(* IEC 61131-3 sources: llm-plc-st-eval/codesys (part 2) *)

(* ---- PRG_Test_I2.st ---- *)
(*
    BANCO DE PRUEBA AUTOVERIFICABLE — Tarea I2 (FSM de llenado multietapa)
    ---------------------------------------------------------------------------
    Reposo -> llenado -> mezcla 60 s -> descarga -> reposo. El paro debe llevar
    a estado seguro (todas las salidas desactivadas) desde CUALQUIER etapa y
    devolver el proceso a reposo.

    USO: crear este PROGRAM junto al FUNCTION_BLOCK de la respuesta a evaluar y
    ejecutar en modo Simulacion. Al terminar, leer 'veredicto': 1 = supera,
    2 = falla.

    ---------------------------------------------------------------------------
    CORRECCION DEL 2026-09-09 (enmienda 10). Validado con validar_harness_I2.py.
    La version anterior tenia dos fallos:

    FALLO 1 — el paso de "antes de los 60 s" REPROBABA a la implementacion
    correcta en los tres ciclos de tarea. Esperaba 59 800 ms contando desde el
    inicio de ese paso, pero la mezcla no arranca ahi: arranca ~200 ms antes,
    en el paso anterior, en cuanto el bloque ve nivelAlto. El margen resultante
    era nulo y la evaluacion caia justo en el instante en que la mezcla
    termina, de modo que se observaba ya la descarga. Es el mismo error que la
    enmienda 5 corrigio en I4: una ventana calculada como si la fase empezara
    en el limite del paso, cuando empieza antes.

    FALLO 2 — el ultimo paso, etiquetado "paro en mezcla", NUNCA llegaba a la
    mezcla. Aplicaba nivelAlto y btnParo en el MISMO paso, asi que el paro
    alcanzaba al bloque todavia en llenado: era un duplicado del paso anterior.
    Verificado: una implementacion cuyo paro funciona en llenado pero no
    durante la mezcla obtenia el mismo resultado que la correcta. El paro en
    dos fases que este banco dice comprobar solo se comprobaba en una.

    La correccion de tiempos de este documento ya lo insinuaba al estimar I2 en
    ~90 s "porque el paro se prueba en dos fases distintas, cada una exige
    volver a entrar en la fase": la secuencia real duraba 61,9 s porque esa
    segunda entrada nunca se hacia.

    Correcciones: la ventana de la mezcla pasa a tener margen explicito y
    simetrico de 0,5 s a cada lado de los 60 s; y entrar en la mezcla y aplicar
    el paro pasan a ser dos pasos separados, de modo que el paro alcance al
    bloque realmente mezclando. Se anade ademas un paso final que comprueba que
    tras el paro el proceso permanece en reposo y no rearranca solo.
*)

PROGRAM PRG_Test_I2
VAR CONSTANT
    ULTIMO_PASO : INT := 11;          (* 12 pasos: indices 0..11 *)
END_VAR
VAR
    (* --- Bloque bajo prueba: sustituir por la respuesta a evaluar --- *)
    fb : FB_Llenado;

    (* --- Entradas manipuladas por el banco --- *)
    nivelAlto : BOOL;
    nivelBajo : BOOL;
    btnInicio : BOOL;
    btnParo   : BOOL;

    (* --- Control de la secuencia --- *)
    evL, evM, evD : BOOL;
    paso       : INT := 0;
    tEspera    : TIME;
    tPaso      : TON;
    pulsoReset : BOOL;
    finalizado : BOOL;

    (* --- Resultados: 0 = pendiente, 1 = pasa, 2 = falla --- *)
    resultado : ARRAY[0..11] OF INT;
    nPasan    : INT;
    veredicto : INT := 0;
    i         : INT;
END_VAR

(* 1. Definicion del paso en curso *)
IF NOT finalizado THEN
    CASE paso OF
        0:  (* Reposo *)
            nivelAlto := FALSE; nivelBajo := FALSE;
            btnInicio := FALSE; btnParo := FALSE;
            tEspera := T#200MS; evL := FALSE; evM := FALSE; evD := FALSE;
        1:  (* Arranque: abre la valvula de llenado *)
            btnInicio := TRUE;
            tEspera := T#200MS; evL := TRUE;  evM := FALSE; evD := FALSE;
        2:  (* Nivel alto: entra en mezcla. La mezcla arranca AQUI, no en el
               paso siguiente; de ahi el margen explicito del paso 3. *)
            btnInicio := FALSE; nivelAlto := TRUE;
            tEspera := T#1S;    evL := FALSE; evM := TRUE;  evD := FALSE;
        3:  (* ~59,5 s de mezcla acumulados: aun NO debe haber terminado *)
            tEspera := T#58500MS; evM := TRUE;
        4:  (* ~60,5 s acumulados: ya debe estar descargando *)
            tEspera := T#1S;    evL := FALSE; evM := FALSE; evD := TRUE;
        5:  (* Nivel bajo: vuelve a reposo *)
            nivelBajo := TRUE;
            tEspera := T#200MS; evL := FALSE; evM := FALSE; evD := FALSE;

        (* --- Paro en la fase de LLENADO --- *)
        6:  (* Nuevo ciclo *)
            nivelAlto := FALSE; nivelBajo := FALSE; btnInicio := TRUE;
            tEspera := T#200MS; evL := TRUE;  evM := FALSE; evD := FALSE;
        7:  (* Paro estando en llenado: estado seguro *)
            btnInicio := FALSE; btnParo := TRUE;
            tEspera := T#200MS; evL := FALSE; evM := FALSE; evD := FALSE;

        (* --- Paro en la fase de MEZCLA (enmienda 10): entrar en la mezcla y
               aplicar el paro son DOS pasos distintos, para que el paro
               alcance al bloque realmente mezclando --- *)
        8:  (* Rearranca tras el paro *)
            btnParo := FALSE; btnInicio := TRUE;
            tEspera := T#200MS; evL := TRUE;  evM := FALSE; evD := FALSE;
        9:  (* Entra en mezcla y se deja mezclando *)
            btnInicio := FALSE; nivelAlto := TRUE;
            tEspera := T#500MS; evL := FALSE; evM := TRUE;  evD := FALSE;
        10: (* Paro ESTANDO EN MEZCLA: estado seguro *)
            btnParo := TRUE;
            tEspera := T#200MS; evL := FALSE; evM := FALSE; evD := FALSE;
        11: (* Tras el paro debe permanecer en reposo, sin rearrancar solo *)
            btnParo := FALSE; nivelAlto := FALSE;
            tEspera := T#200MS; evL := FALSE; evM := FALSE; evD := FALSE;
    END_CASE
END_IF

(* 2. Temporizador de asentamiento del paso *)
tPaso(IN := NOT pulsoReset, PT := tEspera);
pulsoReset := FALSE;

(* 3. Llamada al bloque bajo prueba *)
fb(nivelAlto := nivelAlto, nivelBajo := nivelBajo,
   btnInicio := btnInicio, btnParo := btnParo);

(* 4. Evaluacion al vencer el asentamiento *)
IF tPaso.Q AND NOT finalizado THEN
    IF fb.vLlenado = evL AND fb.motorMezcla = evM AND fb.vDescarga = evD THEN
        resultado[paso] := 1;
    ELSE
        resultado[paso] := 2;
    END_IF

    pulsoReset := TRUE;

    IF paso < ULTIMO_PASO THEN
        paso := paso + 1;
    ELSE
        finalizado := TRUE;
    END_IF
END_IF

(* 5. Veredicto global *)
IF finalizado AND veredicto = 0 THEN
    nPasan := 0;
    FOR i := 0 TO ULTIMO_PASO DO
        IF resultado[i] = 1 THEN
            nPasan := nPasan + 1;
        END_IF
    END_FOR

    IF nPasan = (ULTIMO_PASO + 1) THEN
        veredicto := 1;
    ELSE
        veredicto := 2;
    END_IF
END_IF

(* ---- PRG_Test_I3.st ---- *)
(*
    BANCO DE PRUEBA AUTOVERIFICABLE — Tarea I3 (gestion de alarmas con prioridad)
    ---------------------------------------------------------------------------
    Tres alarmas con prioridad (alm1 alta, alm2 media, alm3 baja). Cualquiera
    activa enciende la sirena. codigoAlm reporta la de mayor prioridad presente
    (0 si no hay). Cada alarma queda RETENIDA aunque su causa desaparezca hasta
    que se reconozca individualmente, y el reconocimiento SOLO tiene efecto si
    la causa ya desaparecio.

    USO: crear este PROGRAM junto al FUNCTION_BLOCK de la respuesta a evaluar y
    ejecutar en modo Simulacion. Al terminar, leer 'veredicto': 1 = supera,
    2 = falla.

    ---------------------------------------------------------------------------
    CORRECCION DEL 2026-09-09 (enmienda 12). Validado con validar_harness_I3.py.
    La version anterior daba veredicto 1 a una implementacion cuyo ACK borraba
    la alarma AUNQUE la causa siguiera presente, que es la violacion directa de
    la regla central del enunciado. Los nueve pasos daban exactamente el mismo
    resultado que con la implementacion correcta.

    Causa: en toda la secuencia no habia un solo instante en que una entrada
    ackN estuviera activa a la vez que su almN. Los reconocimientos se
    aplicaban siempre con la causa ya retirada, de modo que la mitad de la
    regla ("no debe borrar con la causa presente") no se ejercitaba nunca.

    Es notable porque ENMIENDAS_HARNESSES.md ya aprobaba explicitamente ese
    paso en su lista: "I3: ACK con la causa todavia presente (no debe borrar) y
    ACK tras retirarla (si debe)". El paso estaba aprobado en el documento pero
    no implementado en el banco.

    Correccion: se anade el paso 2, que aplica ack3 con alm3 todavia activa y
    exige que la alarma NO se borre. La secuencia pasa de 9 a 10 pasos.
*)

PROGRAM PRG_Test_I3
VAR CONSTANT
    ULTIMO_PASO    : INT  := 9;       (* 10 pasos: indices 0..9 *)
    T_ASENTAMIENTO : TIME := T#150MS;
END_VAR
VAR
    (* --- Bloque bajo prueba: sustituir por la respuesta a evaluar --- *)
    fb : FB_Alarmas;

    (* --- Entradas manipuladas por el banco --- *)
    alm1, alm2, alm3 : BOOL;
    ack1, ack2, ack3 : BOOL;

    (* --- Control de la secuencia --- *)
    espSirena  : BOOL;
    espCodigo  : INT;
    paso       : INT := 0;
    tPaso      : TON;
    pulsoReset : BOOL;
    finalizado : BOOL;

    (* --- Resultados: 0 = pendiente, 1 = pasa, 2 = falla --- *)
    resultado : ARRAY[0..9] OF INT;
    nPasan    : INT;
    veredicto : INT := 0;
    i         : INT;
END_VAR

(* 1. Temporizador de asentamiento entre pasos *)
tPaso(IN := NOT pulsoReset, PT := T_ASENTAMIENTO);
pulsoReset := FALSE;

(* 2. Aplicacion de entradas y valores esperados. Solo se asigna lo que cada
      paso cambia: las demas entradas conservan su valor. *)
IF NOT finalizado THEN
    CASE paso OF
        0:  (* Reposo: sin alarmas, con los ACK activos (no deben hacer nada) *)
            alm1 := FALSE; alm2 := FALSE; alm3 := FALSE;
            ack1 := TRUE;  ack2 := TRUE;  ack3 := TRUE;
            espSirena := FALSE; espCodigo := 0;
        1:  (* Alarma baja activa *)
            ack1 := FALSE; ack2 := FALSE; ack3 := FALSE;
            alm3 := TRUE;
            espSirena := TRUE;  espCodigo := 3;
        2:  (* ACK CON LA CAUSA TODAVIA PRESENTE: no debe borrar (enmienda 12) *)
            ack3 := TRUE;
            espSirena := TRUE;  espCodigo := 3;
        3:  (* Se retira la causa y se suelta el ACK: sigue retenida *)
            alm3 := FALSE; ack3 := FALSE;
            espSirena := TRUE;  espCodigo := 3;
        4:  (* ACK con la causa ya retirada: ahora si debe borrar *)
            ack3 := TRUE;
            espSirena := FALSE; espCodigo := 0;
        5:  (* Dos alarmas: domina la de mayor prioridad de las presentes *)
            ack3 := FALSE; alm2 := TRUE; alm3 := TRUE;
            espSirena := TRUE;  espCodigo := 2;
        6:  (* Entra la de prioridad alta *)
            alm1 := TRUE;
            espSirena := TRUE;  espCodigo := 1;
        7:  (* Se retira y reconoce la alta: queda la media *)
            alm1 := FALSE; ack1 := TRUE;
            espSirena := TRUE;  espCodigo := 2;
        8:  (* Se retira y reconoce la media: queda la baja *)
            alm2 := FALSE; ack2 := TRUE;
            espSirena := TRUE;  espCodigo := 3;
        9:  (* Se retira y reconoce la baja: todo en reposo *)
            alm3 := FALSE; ack3 := TRUE;
            espSirena := FALSE; espCodigo := 0;
    END_CASE
END_IF

(* 3. Llamada al bloque bajo prueba *)
fb(alm1 := alm1, alm2 := alm2, alm3 := alm3,
   ack1 := ack1, ack2 := ack2, ack3 := ack3);

(* 4. Evaluacion al vencer el asentamiento *)
IF tPaso.Q AND NOT finalizado THEN
    IF fb.sirena = espSirena AND fb.codigoAlm = espCodigo THEN
        resultado[paso] := 1;
    ELSE
        resultado[paso] := 2;
    END_IF

    pulsoReset := TRUE;

    IF paso < ULTIMO_PASO THEN
        paso := paso + 1;
    ELSE
        finalizado := TRUE;
    END_IF
END_IF

(* 5. Veredicto global *)
IF finalizado AND veredicto = 0 THEN
    nPasan := 0;
    FOR i := 0 TO ULTIMO_PASO DO
        IF resultado[i] = 1 THEN
            nPasan := nPasan + 1;
        END_IF
    END_FOR

    IF nPasan = (ULTIMO_PASO + 1) THEN
        veredicto := 1;
    ELSE
        veredicto := 2;
    END_IF
END_IF

(* ---- PRG_Test_I4.st ---- *)
(*
    BANCO DE PRUEBA AUTOVERIFICABLE — Tarea I4 (arranque estrella-triangulo)
    ---------------------------------------------------------------------------
    Aplica la enmienda 2 de ENMIENDAS_HARNESSES.md: DOS verificaciones
    independientes, porque una transicion con 0 ms de tiempo muerto no produce
    ningun scan con kY AND kD y por tanto la bandera de interlock por si sola
    no la detecta.
      1. Seguridad (continua y enclavada): si en cualquier scan kY AND kD, la
         bandera 'interlock' queda en TRUE hasta el final del banco.
      2. Tiempo muerto (medido): se cronometra el intervalo entre la caida de
         kY y la subida de kD y se exige que alcance el minimo.

    Ciclo de MainTask: 4 a 10 ms (enmienda 3). El umbral del tiempo muerto
    absorbe un ciclo de cuantizacion del scan.

    USO: crear este PROGRAM junto al FUNCTION_BLOCK de la respuesta a evaluar y
    ejecutar en modo Simulacion. Al terminar, leer 'veredicto': 1 = supera,
    2 = falla. 'resultado' indica el paso; 'interlock' y 'duracionMuerto' se
    registran aparte porque una violacion de seguridad es cualitativamente
    distinta de un fallo funcional (enmienda 4).

    ---------------------------------------------------------------------------
    CORRECCION DEL 2026-09-09 (enmienda 5). La version anterior tenia tres
    fallos, verificados por simulacion con validar_harness_I4.py:

      1. El paso 2 exigia NOT kD a los 8,3 s, cuando una implementacion
         correcta ya tiene el triangulo dentro desde los 8,1 s. Reprobaba al
         100 % de las implementaciones validas. Era un residuo del enfoque de
         muestreo que la enmienda 2 habia descartado.
      2. La medida reiniciaba su temporizador con un ciclo de retraso, de modo
         que contaba de menos alrededor de un scan: un tiempo muerto correcto
         de 100 ms se media como 96 ms con ciclo de 4 ms y 80 ms con 20 ms, y
         se comparaba contra un umbral estricto de 100 ms.
      3. Si kY caia y kD subia en el MISMO scan, ambas condiciones se cumplian
         en el mismo ciclo, la medida leia un valor viejo del cronometro y
         registraba 8 208 ms: daba por bueno el defecto de 0 ms de tiempo
         muerto, que es exactamente el que la enmienda 2 persigue.

    La medida pasa a hacerse por DIFERENCIA de dos lecturas de un cronometro
    libre que nunca se reinicia. Eso elimina el retraso de un ciclo y hace que
    el caso simultaneo mida 0 ms por construccion, sin necesidad de un caso
    especial. El paso 2 pasa a comprobar que la transicion se completo, y el
    instante exacto queda a cargo de la medida en el paso 3.
*)

PROGRAM PRG_Test_I4
VAR CONSTANT
    ULTIMO_PASO   : INT  := 5;
    T_MUERTO_MIN  : TIME := T#90MS;   (* 100 ms del enunciado menos un ciclo de
                                         MainTask: la cuantizacion del scan es
                                         inevitable y se declara en la metodologia *)
    T_CRONO       : TIME := T#100S;   (* cronometro libre: nunca se reinicia *)
END_VAR
VAR
    (* --- Bloque bajo prueba: sustituir por la respuesta a evaluar --- *)
    fb : FB_EstrellaTriangulo;

    (* --- Entradas manipuladas por el banco --- *)
    btnMarcha : BOOL;
    btnParo   : BOOL;

    (* --- Control de la secuencia --- *)
    paso       : INT := 0;
    tEspera    : TIME;
    tPaso      : TON;
    pulsoReset : BOOL;
    finalizado : BOOL;

    (* --- Verificacion 1: seguridad continua y enclavada (enmiendas 2 y 4) --- *)
    interlock : BOOL;

    (* --- Verificacion 2: medida del tiempo muerto (enmienda 2) --- *)
    tCrono         : TON;
    prevY, prevD   : BOOL;
    midiendo       : BOOL;
    etCaidaY       : TIME;
    duracionMuerto : TIME;
    muertoOK       : BOOL;

    (* --- Resultados: 0 = pendiente, 1 = pasa, 2 = falla --- *)
    resultado : ARRAY[0..5] OF INT;
    nPasan    : INT;
    veredicto : INT := 0;
    i         : INT;
END_VAR

(* 1. Definicion del paso en curso. Va antes del temporizador porque tEspera
      lo alimenta. Solo se asigna lo que cada paso cambia. *)
IF NOT finalizado THEN
    CASE paso OF
        0:  (* Reposo *)
            btnMarcha := FALSE; btnParo := FALSE;
            tEspera   := T#200MS;
        1:  (* Fase estrella: se evalua antes de los 8 s de transicion *)
            btnMarcha := TRUE;
            tEspera   := T#7800MS;
        2:  (* Ya pasada la transicion: debe estar en triangulo *)
            tEspera   := T#500MS;
        3:  (* Confirmacion del veredicto de tiempo muerto *)
            tEspera   := T#300MS;
        4:  (* Paro en cualquier momento: todo a reposo *)
            btnMarcha := FALSE; btnParo := TRUE;
            tEspera   := T#200MS;
        5:  (* Rearranque: debe volver a estrella, no saltar a triangulo *)
            btnParo := FALSE; btnMarcha := TRUE;
            tEspera := T#200MS;
    END_CASE
END_IF

(* 2. Temporizadores del banco *)
tPaso(IN := NOT pulsoReset, PT := tEspera);
tCrono(IN := TRUE, PT := T_CRONO);
pulsoReset := FALSE;

(* 3. Llamada al bloque bajo prueba *)
fb(btnMarcha := btnMarcha, btnParo := btnParo);

(* 4. Verificacion 1 — seguridad: se evalua en CADA scan y queda enclavada *)
IF fb.kY AND fb.kD THEN
    interlock := TRUE;
END_IF

(* 5. Verificacion 2 — tiempo muerto por diferencia de dos lecturas del
      cronometro libre. Si kY cae y kD sube en el mismo scan, ambas ramas se
      ejecutan en ese ciclo y la diferencia vale 0: el defecto queda detectado
      sin necesidad de un caso especial. *)
IF prevY AND NOT fb.kY THEN
    etCaidaY := tCrono.ET;
    midiendo := TRUE;
END_IF

IF midiendo AND fb.kD AND NOT prevD THEN
    duracionMuerto := tCrono.ET - etCaidaY;
    IF duracionMuerto >= T_MUERTO_MIN THEN
        muertoOK := TRUE;
    END_IF
    midiendo := FALSE;
END_IF

prevY := fb.kY;
prevD := fb.kD;

(* 6. Evaluacion al vencer el asentamiento del paso *)
IF tPaso.Q AND NOT finalizado THEN
    IF    (paso = 0 AND NOT fb.kM AND NOT fb.kY AND NOT fb.kD)
       OR (paso = 1 AND fb.kM AND fb.kY AND NOT fb.kD)
       OR (paso = 2 AND fb.kM AND NOT fb.kY AND fb.kD)
       OR (paso = 3 AND fb.kM AND NOT fb.kY AND fb.kD AND muertoOK)
       OR (paso = 4 AND NOT fb.kM AND NOT fb.kY AND NOT fb.kD)
       OR (paso = 5 AND fb.kM AND fb.kY AND NOT fb.kD)
    THEN
        resultado[paso] := 1;
    ELSE
        resultado[paso] := 2;
    END_IF

    pulsoReset := TRUE;

    IF paso < ULTIMO_PASO THEN
        paso := paso + 1;
    ELSE
        finalizado := TRUE;
    END_IF
END_IF

(* 7. Veredicto global: exige superar todos los pasos Y no haber violado
      nunca el interlock (enmienda 4) *)
IF finalizado AND veredicto = 0 THEN
    nPasan := 0;
    FOR i := 0 TO ULTIMO_PASO DO
        IF resultado[i] = 1 THEN
            nPasan := nPasan + 1;
        END_IF
    END_FOR

    IF nPasan = (ULTIMO_PASO + 1) AND NOT interlock THEN
        veredicto := 1;
    ELSE
        veredicto := 2;
    END_IF
END_IF

(* ---- PRG_Test_I5.st ---- *)
(*
    BANCO DE PRUEBA AUTOVERIFICABLE — Tarea I5 (banda clasificadora)
    ---------------------------------------------------------------------------
    La banda funciona siempre. Cada flanco de sensorPresencia cuenta una pieza;
    si sensorAltura esta activo en ese instante la pieza es alta y debe
    desviarse: el piston se activa durante 1 s, comenzando 2 s despues de la
    deteccion. Se cuentan altas y bajas por separado.

    USO: crear este PROGRAM junto al FUNCTION_BLOCK de la respuesta a evaluar y
    ejecutar en modo Simulacion. Al terminar, leer 'veredicto': 1 = supera,
    2 = falla.

    ---------------------------------------------------------------------------
    CORRECCION DEL 2026-09-09 (enmienda 11). Validado con validar_harness_I5.py.
    La version anterior REPROBABA a la implementacion correcta en los tres
    ciclos de tarea.

    Causa: el paso que decia comprobar "antes de 2 s" esperaba 1800 ms contando
    desde su propio inicio, pero la deteccion de la pieza alta ocurre 200 ms
    antes, en el paso anterior. El tiempo efectivo desde la deteccion era por
    tanto de 2000 ms exactos, es decir justo el instante en que el piston se
    activa, y la evaluacion lo encontraba ya activado.

    Es el tercer caso del mismo error, tras I4 (enmienda 5) e I2 (enmienda 10):
    una ventana calculada como si la fase empezara en el limite del paso,
    cuando en realidad empieza antes. Conviene enunciarlo como regla: el
    tiempo de una ventana se cuenta desde el evento que la origina, no desde
    el paso en que se escribe.

    Correccion: las tres ventanas del desvio se recalculan con margen explicito
    de 0,3 s a 0,5 s respecto a los flancos del pulso, tomando como origen la
    deteccion real. Con la secuencia corregida se discriminan un retardo de
    1,5 s, la ausencia de retardo, un pulso de 2 s y el desvio indebido de las
    piezas bajas.

    Cronologia (t = 0 en el arranque del banco; deteccion de la pieza alta en
    t = 0,7 s; pulso correcto de 2,7 s a 3,7 s):
        paso 4 evalua en t = 2,4 s  -> 0,3 s ANTES de que el piston se active
        paso 5 evalua en t = 3,2 s  -> dentro del pulso, a 0,5 s de cada flanco
        paso 6 evalua en t = 4,0 s  -> 0,3 s DESPUES de que el piston se apague
*)

PROGRAM PRG_Test_I5
VAR CONSTANT
    ULTIMO_PASO : INT := 6;
END_VAR
VAR
    (* --- Bloque bajo prueba: sustituir por la respuesta a evaluar --- *)
    fb : FB_Clasificadora;

    (* --- Entradas manipuladas por el banco --- *)
    sensorPresencia : BOOL;
    sensorAltura    : BOOL;

    (* --- Control de la secuencia --- *)
    espBanda, espPiston : BOOL;
    espAltas, espBajas  : INT;
    paso       : INT := 0;
    tEspera    : TIME;
    tPaso      : TON;
    pulsoReset : BOOL;
    finalizado : BOOL;

    (* --- Resultados: 0 = pendiente, 1 = pasa, 2 = falla --- *)
    resultado : ARRAY[0..6] OF INT;
    nPasan    : INT;
    veredicto : INT := 0;
    i         : INT;
END_VAR

(* 1. Definicion del paso en curso *)
IF NOT finalizado THEN
    CASE paso OF
        0:  (* Reposo: la banda debe estar en marcha desde el principio *)
            sensorPresencia := FALSE; sensorAltura := FALSE;
            tEspera := T#200MS;
            espBanda := TRUE; espPiston := FALSE; espAltas := 0; espBajas := 0;
        1:  (* Pieza baja con presencia SOSTENIDA: debe contar una sola vez *)
            sensorPresencia := TRUE; sensorAltura := FALSE;
            tEspera := T#300MS;
            espBanda := TRUE; espPiston := FALSE; espAltas := 0; espBajas := 1;
        2:  (* Se retira la pieza baja *)
            sensorPresencia := FALSE;
            tEspera := T#200MS;
            espBanda := TRUE; espPiston := FALSE; espAltas := 0; espBajas := 1;
        3:  (* Pieza ALTA: aqui empieza a contar el retardo de 2 s del desvio *)
            sensorPresencia := TRUE; sensorAltura := TRUE;
            tEspera := T#200MS;
            espBanda := TRUE; espPiston := FALSE; espAltas := 1; espBajas := 1;

        (* --- Ventanas del desvio, con origen en la deteccion (enmienda 11) --- *)
        4:  (* t = 2,4 s: 0,3 s antes de que el piston deba activarse *)
            sensorPresencia := FALSE; sensorAltura := FALSE;
            tEspera := T#1500MS;
            espBanda := TRUE; espPiston := FALSE; espAltas := 1; espBajas := 1;
        5:  (* t = 3,2 s: dentro del pulso, a 0,5 s de cada flanco *)
            tEspera := T#800MS;
            espBanda := TRUE; espPiston := TRUE;  espAltas := 1; espBajas := 1;
        6:  (* t = 4,0 s: 0,3 s despues de que el piston deba apagarse *)
            tEspera := T#800MS;
            espBanda := TRUE; espPiston := FALSE; espAltas := 1; espBajas := 1;
    END_CASE
END_IF

(* 2. Temporizador de asentamiento del paso *)
tPaso(IN := NOT pulsoReset, PT := tEspera);
pulsoReset := FALSE;

(* 3. Llamada al bloque bajo prueba *)
fb(sensorPresencia := sensorPresencia, sensorAltura := sensorAltura);

(* 4. Evaluacion al vencer el asentamiento *)
IF tPaso.Q AND NOT finalizado THEN
    IF     fb.banda   = espBanda
       AND fb.piston  = espPiston
       AND fb.nAltas  = espAltas
       AND fb.nBajas  = espBajas
    THEN
        resultado[paso] := 1;
    ELSE
        resultado[paso] := 2;
    END_IF

    pulsoReset := TRUE;

    IF paso < ULTIMO_PASO THEN
        paso := paso + 1;
    ELSE
        finalizado := TRUE;
    END_IF
END_IF

(* 5. Veredicto global *)
IF finalizado AND veredicto = 0 THEN
    nPasan := 0;
    FOR i := 0 TO ULTIMO_PASO DO
        IF resultado[i] = 1 THEN
            nPasan := nPasan + 1;
        END_IF
    END_FOR

    IF nPasan = (ULTIMO_PASO + 1) THEN
        veredicto := 1;
    ELSE
        veredicto := 2;
    END_IF
END_IF

(* ---- PRG_Test_I6.st ---- *)
(*
    BANCO DE PRUEBA AUTOVERIFICABLE — Tarea I6 (escalado analogico con histeresis)
    ---------------------------------------------------------------------------
    rawTemp de 0 a 27648 se escala a tempC de 0.0 a 100.0 grados. El enfriador
    se activa cuando tempC alcanza 80.0 y se desactiva cuando desciende a 75.0,
    conservando su estado entre ambos umbrales. Si rawTemp queda fuera del
    rango se activa almSensor Y SE DESACTIVA EL ENFRIADOR.

    Se comprueba la histeresis en LOS DOS SENTIDOS: conserva el estado ON al
    bajar dentro de la banda y conserva el estado OFF al subir dentro de ella.

    USO: crear este PROGRAM junto al FUNCTION_BLOCK de la respuesta a evaluar y
    ejecutar en modo Simulacion. Al terminar, leer 'veredicto': 1 = supera,
    2 = falla.

    ---------------------------------------------------------------------------
    CORRECCION DEL 2026-09-09 (enmienda 13). Validado con validar_harness_I6.py.
    La version anterior daba veredicto 1 a una implementacion que activaba la
    alarma pero NO desactivaba el enfriador, incumpliendo la ultima frase del
    enunciado.

    Causa: los dos pasos de fuera de rango estaban al final de la secuencia,
    cuando el enfriador ya llevaba tres pasos apagado. La condicion "y se
    desactiva el enfriador" se evaluaba sobre una salida que ya estaba en el
    valor esperado, de modo que la implementacion defectuosa y la correcta
    daban el mismo resultado. Para observar que la alarma APAGA el enfriador
    hay que provocarla con el enfriador ENCENDIDO.

    Es el mismo patron de cobertura de las enmiendas 7, 9, 10 y 12: el banco no
    llegaba al estado en el que el defecto se manifiesta.

    Correccion: el primer paso de fuera de rango se adelanta y pasa a aplicarse
    justo despues de la banda de histeresis con el enfriador encendido. La
    secuencia conserva los ocho pasos y sigue cubriendo los dos sentidos de la
    histeresis y los dos limites del rango.
*)

PROGRAM PRG_Test_I6
VAR CONSTANT
    ULTIMO_PASO    : INT  := 7;
    T_ASENTAMIENTO : TIME := T#100MS;
    RAW_MAX        : INT  := 27648;
END_VAR
VAR
    (* --- Bloque bajo prueba: sustituir por la respuesta a evaluar --- *)
    fb : FB_Temperatura;

    (* --- Entrada manipulada por el banco --- *)
    rawTemp : INT;

    (* --- Control de la secuencia --- *)
    espTemp    : REAL;
    espFrio    : BOOL;
    espAlarma  : BOOL;
    compTemp   : BOOL;                (* FALSE fuera de rango: tempC indefinida *)
    paso       : INT := 0;
    tPaso      : TON;
    pulsoReset : BOOL;
    finalizado : BOOL;

    (* --- Resultados: 0 = pendiente, 1 = pasa, 2 = falla --- *)
    resultado : ARRAY[0..7] OF INT;
    nPasan    : INT;
    veredicto : INT := 0;
    i         : INT;
END_VAR

(* 1. Temporizador de asentamiento entre pasos *)
tPaso(IN := NOT pulsoReset, PT := T_ASENTAMIENTO);
pulsoReset := FALSE;

(* 2. Definicion del paso en curso *)
IF NOT finalizado THEN
    CASE paso OF
        0:  (* Punto medio del rango *)
            rawTemp := 13824; espTemp := 50.0;
            espFrio := FALSE; espAlarma := FALSE; compTemp := TRUE;
        1:  (* Umbral superior: el enfriador debe activarse *)
            rawTemp := 22119; espTemp := 80.0;
            espFrio := TRUE;  espAlarma := FALSE; compTemp := TRUE;
        2:  (* Dentro de la banda bajando: debe CONSERVAR el estado ON *)
            rawTemp := 21289; espTemp := 77.0;
            espFrio := TRUE;  espAlarma := FALSE; compTemp := TRUE;
        3:  (* Fuera de rango CON EL ENFRIADOR ENCENDIDO (enmienda 13):
               la alarma debe activarse y el enfriador debe apagarse *)
            rawTemp := 27649; espTemp := 0.0;
            espFrio := FALSE; espAlarma := TRUE;  compTemp := FALSE;
        4:  (* Vuelve al rango en el umbral inferior: enfriador apagado *)
            rawTemp := 20736; espTemp := 75.0;
            espFrio := FALSE; espAlarma := FALSE; compTemp := TRUE;
        5:  (* Dentro de la banda subiendo: debe CONSERVAR el estado OFF *)
            rawTemp := 21289; espTemp := 77.0;
            espFrio := FALSE; espAlarma := FALSE; compTemp := TRUE;
        6:  (* Fuera de rango por el limite inferior *)
            rawTemp := -1;    espTemp := 0.0;
            espFrio := FALSE; espAlarma := TRUE;  compTemp := FALSE;
        7:  (* Vuelve al rango: la alarma debe desactivarse *)
            rawTemp := 0;     espTemp := 0.0;
            espFrio := FALSE; espAlarma := FALSE; compTemp := TRUE;
    END_CASE
END_IF

(* 3. Llamada al bloque bajo prueba *)
fb(rawTemp := rawTemp);

(* 4. Evaluacion al vencer el asentamiento. tempC solo se comprueba dentro
      del rango: fuera de el su valor no esta definido por el enunciado. *)
IF tPaso.Q AND NOT finalizado THEN
    IF     fb.enfriador = espFrio
       AND fb.almSensor = espAlarma
       AND ((NOT compTemp)
            OR ((fb.tempC > espTemp - 0.1) AND (fb.tempC < espTemp + 0.1)))
    THEN
        resultado[paso] := 1;
    ELSE
        resultado[paso] := 2;
    END_IF

    pulsoReset := TRUE;

    IF paso < ULTIMO_PASO THEN
        paso := paso + 1;
    ELSE
        finalizado := TRUE;
    END_IF
END_IF

(* 5. Veredicto global *)
IF finalizado AND veredicto = 0 THEN
    nPasan := 0;
    FOR i := 0 TO ULTIMO_PASO DO
        IF resultado[i] = 1 THEN
            nPasan := nPasan + 1;
        END_IF
    END_FOR

    IF nPasan = (ULTIMO_PASO + 1) THEN
        veredicto := 1;
    ELSE
        veredicto := 2;
    END_IF
END_IF

(* ---- PRG_Test_I7.st ---- *)
(*
    BANCO DE PRUEBA AUTOVERIFICABLE - Tarea I7 (FB_Duplex: bombas duplex con alternancia)
    ---------------------------------------------------------------------------
    Validado en codesys/validar_harness_I7.py: 10 implementaciones (la correcta,
    el FB de referencia del prompt de C4 y 8 defectuosas), ciclos de 4, 10 y 20 ms.
    La tabla de pasos se genera desde el validador para que ambos coincidan.

    Paso (demanda, falla1, falla2) -> (bomba1, bomba2, almFalla)   principal
  0  (F,F,F) -> (F,F,F)                                          -
  1  (T,F,F) -> (T,F,F)   primera demanda                        b1
  2  (F,F,F) -> (F,F,F)
  3  (T,F,F) -> (F,T,F)   alterna                                b2
  4  (F,F,F) -> (F,F,F)
  5  (T,F,F) -> (T,F,F)   alterna de nuevo                       b1
  6  (T,T,F) -> (F,T,T)   falla de la principal: respaldo        b1
  7  (T,F,F) -> (T,F,F)   vuelve la principal                    b1
  8  (T,F,T) -> (T,F,F)   falla SOLO del respaldo: sin alarma    b1
  9  (T,T,T) -> (F,F,T)   ambas con falla                        b1
 10  (F,T,T) -> (F,F,F)   sin demanda: sin alarma aunque haya fallas
 11  (T,F,F) -> (F,T,F)   cuarta demanda                         b2
 12  (T,F,T) -> (T,F,T)   falla de la principal b2: respaldo b1  b2
 13  (F,F,F) -> (F,F,F)
*)
PROGRAM PRG_Test_I7
VAR CONSTANT
    ULTIMO_PASO : INT  := 13;
    T_PASO      : TIME := T#100MS;
END_VAR
VAR
    fb : FB_Duplex;                 (* bloque bajo prueba *)
    demanda, falla1, falla2 : BOOL;
    e1, e2, eAlm : BOOL;            (* esperados: bomba1, bomba2, almFalla *)

    paso       : INT := 0;
    tPaso      : TON;
    pulsoReset : BOOL;
    finalizado : BOOL;

    resultado : ARRAY[0..13] OF INT;
    nPasan    : INT;
    veredicto : INT := 0;
    i         : INT;
END_VAR

(* 1. Entradas y salidas esperadas del paso *)
IF NOT finalizado THEN
    CASE paso OF
        0: demanda := FALSE; falla1 := FALSE; falla2 := FALSE;
            e1 := FALSE; e2 := FALSE; eAlm := FALSE;
        1: demanda := TRUE; falla1 := FALSE; falla2 := FALSE;
            e1 := TRUE; e2 := FALSE; eAlm := FALSE;
        2: demanda := FALSE; falla1 := FALSE; falla2 := FALSE;
            e1 := FALSE; e2 := FALSE; eAlm := FALSE;
        3: demanda := TRUE; falla1 := FALSE; falla2 := FALSE;
            e1 := FALSE; e2 := TRUE; eAlm := FALSE;
        4: demanda := FALSE; falla1 := FALSE; falla2 := FALSE;
            e1 := FALSE; e2 := FALSE; eAlm := FALSE;
        5: demanda := TRUE; falla1 := FALSE; falla2 := FALSE;
            e1 := TRUE; e2 := FALSE; eAlm := FALSE;
        6: demanda := TRUE; falla1 := TRUE; falla2 := FALSE;
            e1 := FALSE; e2 := TRUE; eAlm := TRUE;
        7: demanda := TRUE; falla1 := FALSE; falla2 := FALSE;
            e1 := TRUE; e2 := FALSE; eAlm := FALSE;
        8: demanda := TRUE; falla1 := FALSE; falla2 := TRUE;
            e1 := TRUE; e2 := FALSE; eAlm := FALSE;
        9: demanda := TRUE; falla1 := TRUE; falla2 := TRUE;
            e1 := FALSE; e2 := FALSE; eAlm := TRUE;
        10: demanda := FALSE; falla1 := TRUE; falla2 := TRUE;
            e1 := FALSE; e2 := FALSE; eAlm := FALSE;
        11: demanda := TRUE; falla1 := FALSE; falla2 := FALSE;
            e1 := FALSE; e2 := TRUE; eAlm := FALSE;
        12: demanda := TRUE; falla1 := FALSE; falla2 := TRUE;
            e1 := TRUE; e2 := FALSE; eAlm := TRUE;
        13: demanda := FALSE; falla1 := FALSE; falla2 := FALSE;
            e1 := FALSE; e2 := FALSE; eAlm := FALSE;
    END_CASE
END_IF

(* 2. Asentamiento del paso *)
tPaso(IN := NOT pulsoReset, PT := T_PASO);
pulsoReset := FALSE;

(* 3. Bloque bajo prueba *)
fb(demanda := demanda, falla1 := falla1, falla2 := falla2);

(* 4. Evaluacion *)
IF tPaso.Q AND NOT finalizado THEN
    IF (fb.bomba1 = e1) AND (fb.bomba2 = e2) AND (fb.almFalla = eAlm) THEN
        resultado[paso] := 1;
    ELSE
        resultado[paso] := 2;
    END_IF
    pulsoReset := TRUE;
    IF paso < ULTIMO_PASO THEN
        paso := paso + 1;
    ELSE
        finalizado := TRUE;
    END_IF
END_IF

(* 5. Veredicto global *)
IF finalizado AND veredicto = 0 THEN
    nPasan := 0;
    FOR i := 0 TO ULTIMO_PASO DO
        IF resultado[i] = 1 THEN
            nPasan := nPasan + 1;
        END_IF
    END_FOR
    IF nPasan = (ULTIMO_PASO + 1) THEN
        veredicto := 1;
    ELSE
        veredicto := 2;
    END_IF
END_IF

(* ---- PRG_Test_I8.st ---- *)
(*
    BANCO DE PRUEBA AUTOVERIFICABLE - Tarea I8 (FB_Compresor: permisivos de arranque)
    ---------------------------------------------------------------------------
    Validado en codesys/validar_harness_I8.py: 8 implementaciones (1 correcta y
    7 defectuosas), ciclos de 4, 10 y 20 ms. La tabla de pasos se genera desde
    el validador para que ambos coincidan.

    Paso: entradas (pOil,temp,sinAlm,marcha,paro), duracion -> (comp, causa)
  0 (F,F,F,F,F) 0.2 s -> (F,1)   reposo, faltan todos: reporta el menor
  1 (T,T,T,F,F) 1.0 s -> (F,1)   aceite aun sin 3 s continuos
  2 (T,T,T,F,F) 2.5 s -> (F,0)   permisivos completos: NO arranca solo
  3 (T,T,T,T,F) 0.2 s -> (T,0)   flanco de marcha
  4 (T,T,T,F,F) 0.2 s -> (T,0)   enclavado
  5 (T,F,T,F,F) 0.2 s -> (F,2)   pierde temperatura
  6 (T,T,T,F,F) 0.5 s -> (F,0)   se recupera: sin rearranque automatico
  7 (T,T,T,T,T) 0.2 s -> (F,0)   marcha y paro a la vez: prioridad del paro
  8 (T,T,T,T,F) 0.2 s -> (F,0)   se suelta el paro con marcha sostenida: sin flanco no arranca
  9 (T,T,T,F,F) 0.2 s -> (F,0)
 10 (T,T,T,T,F) 0.2 s -> (T,0)
 11 (T,T,F,F,F) 0.2 s -> (F,3)   alarma
 12 (F,F,F,F,F) 0.2 s -> (F,1)   faltan todos
 13 (T,T,T,T,F) 0.5 s -> (F,1)   pulsa con el aceite aun temporizando (reiniciado)
 14 (T,T,T,T,F) 3.0 s -> (F,0)   llegan los permisivos con marcha sostenida: no arranca
 15 (T,T,T,F,F) 0.2 s -> (F,0)
 16 (T,T,T,T,F) 0.2 s -> (T,0)
 17 (F,T,T,T,F) 0.2 s -> (F,1)   perdida momentanea de aceite: se detiene
 18 (T,T,T,F,F) 0.2 s -> (F,1)   el aceite vuelve pero no lleva 3 s

VIGILANCIA CONTINUA (patron de la enmienda 4, banderas enclavadas): en los pasos
en que comp llega en FALSE y debe seguir en FALSE todo el paso (0,1,2,6,7,8,9,
12,13,14,15,18), un solo scan con comp=TRUE reprueba el paso. Sin ella, la
validacion mostro que "marcha gana al paro" pasaba inadvertido: el compresor
arrancaba UN scan en el paso 7 y se apagaba antes del muestreo.
*)
PROGRAM PRG_Test_I8
VAR CONSTANT
    ULTIMO_PASO : INT := 18;
END_VAR
VAR
    fb : FB_Compresor;              (* bloque bajo prueba *)
    pOilOk, tempOk, sinAlm, btnMarcha, btnParo : BOOL;
    eComp  : BOOL;                  (* esperado *)
    eCausa : INT;

    paso       : INT := 0;
    tEspera    : TIME;
    tPaso      : TON;
    pulsoReset : BOOL;
    finalizado : BOOL;
    vigilado   : BOOL;
    violacion  : BOOL;              (* bandera enclavada del paso *)

    resultado : ARRAY[0..18] OF INT;
    nPasan    : INT;
    veredicto : INT := 0;
    i         : INT;
END_VAR

(* 1. Entradas, duracion y salidas esperadas del paso *)
IF NOT finalizado THEN
    CASE paso OF
        0: pOilOk := FALSE; tempOk := FALSE; sinAlm := FALSE; btnMarcha := FALSE; btnParo := FALSE;
            tEspera := T#200MS; eComp := FALSE; eCausa := 1;
        1: pOilOk := TRUE; tempOk := TRUE; sinAlm := TRUE; btnMarcha := FALSE; btnParo := FALSE;
            tEspera := T#1000MS; eComp := FALSE; eCausa := 1;
        2: pOilOk := TRUE; tempOk := TRUE; sinAlm := TRUE; btnMarcha := FALSE; btnParo := FALSE;
            tEspera := T#2500MS; eComp := FALSE; eCausa := 0;
        3: pOilOk := TRUE; tempOk := TRUE; sinAlm := TRUE; btnMarcha := TRUE; btnParo := FALSE;
            tEspera := T#200MS; eComp := TRUE; eCausa := 0;
        4: pOilOk := TRUE; tempOk := TRUE; sinAlm := TRUE; btnMarcha := FALSE; btnParo := FALSE;
            tEspera := T#200MS; eComp := TRUE; eCausa := 0;
        5: pOilOk := TRUE; tempOk := FALSE; sinAlm := TRUE; btnMarcha := FALSE; btnParo := FALSE;
            tEspera := T#200MS; eComp := FALSE; eCausa := 2;
        6: pOilOk := TRUE; tempOk := TRUE; sinAlm := TRUE; btnMarcha := FALSE; btnParo := FALSE;
            tEspera := T#500MS; eComp := FALSE; eCausa := 0;
        7: pOilOk := TRUE; tempOk := TRUE; sinAlm := TRUE; btnMarcha := TRUE; btnParo := TRUE;
            tEspera := T#200MS; eComp := FALSE; eCausa := 0;
        8: pOilOk := TRUE; tempOk := TRUE; sinAlm := TRUE; btnMarcha := TRUE; btnParo := FALSE;
            tEspera := T#200MS; eComp := FALSE; eCausa := 0;
        9: pOilOk := TRUE; tempOk := TRUE; sinAlm := TRUE; btnMarcha := FALSE; btnParo := FALSE;
            tEspera := T#200MS; eComp := FALSE; eCausa := 0;
        10: pOilOk := TRUE; tempOk := TRUE; sinAlm := TRUE; btnMarcha := TRUE; btnParo := FALSE;
            tEspera := T#200MS; eComp := TRUE; eCausa := 0;
        11: pOilOk := TRUE; tempOk := TRUE; sinAlm := FALSE; btnMarcha := FALSE; btnParo := FALSE;
            tEspera := T#200MS; eComp := FALSE; eCausa := 3;
        12: pOilOk := FALSE; tempOk := FALSE; sinAlm := FALSE; btnMarcha := FALSE; btnParo := FALSE;
            tEspera := T#200MS; eComp := FALSE; eCausa := 1;
        13: pOilOk := TRUE; tempOk := TRUE; sinAlm := TRUE; btnMarcha := TRUE; btnParo := FALSE;
            tEspera := T#500MS; eComp := FALSE; eCausa := 1;
        14: pOilOk := TRUE; tempOk := TRUE; sinAlm := TRUE; btnMarcha := TRUE; btnParo := FALSE;
            tEspera := T#3000MS; eComp := FALSE; eCausa := 0;
        15: pOilOk := TRUE; tempOk := TRUE; sinAlm := TRUE; btnMarcha := FALSE; btnParo := FALSE;
            tEspera := T#200MS; eComp := FALSE; eCausa := 0;
        16: pOilOk := TRUE; tempOk := TRUE; sinAlm := TRUE; btnMarcha := TRUE; btnParo := FALSE;
            tEspera := T#200MS; eComp := TRUE; eCausa := 0;
        17: pOilOk := FALSE; tempOk := TRUE; sinAlm := TRUE; btnMarcha := TRUE; btnParo := FALSE;
            tEspera := T#200MS; eComp := FALSE; eCausa := 1;
        18: pOilOk := TRUE; tempOk := TRUE; sinAlm := TRUE; btnMarcha := FALSE; btnParo := FALSE;
            tEspera := T#200MS; eComp := FALSE; eCausa := 1;
    END_CASE
END_IF

(* 2. Asentamiento del paso *)
tPaso(IN := NOT pulsoReset, PT := tEspera);
pulsoReset := FALSE;

(* 3. Bloque bajo prueba *)
fb(pOilOk := pOilOk, tempOk := tempOk, sinAlm := sinAlm, btnMarcha := btnMarcha, btnParo := btnParo);

(* 4. Vigilancia continua: comp no puede valer TRUE ni un scan en estos pasos *)
CASE paso OF
    0, 1, 2, 6, 7, 8, 9, 12, 13, 14, 15, 18: vigilado := TRUE;
ELSE
    vigilado := FALSE;
END_CASE
IF vigilado AND fb.comp AND NOT finalizado THEN
    violacion := TRUE;
END_IF

(* 5. Evaluacion *)
IF tPaso.Q AND NOT finalizado THEN
    IF (fb.comp = eComp) AND (fb.causaBloqueo = eCausa) AND NOT violacion THEN
        resultado[paso] := 1;
    ELSE
        resultado[paso] := 2;
    END_IF
    violacion := FALSE;
    pulsoReset := TRUE;
    IF paso < ULTIMO_PASO THEN
        paso := paso + 1;
    ELSE
        finalizado := TRUE;
    END_IF
END_IF

(* 6. Veredicto global *)
IF finalizado AND veredicto = 0 THEN
    nPasan := 0;
    FOR i := 0 TO ULTIMO_PASO DO
        IF resultado[i] = 1 THEN
            nPasan := nPasan + 1;
        END_IF
    END_FOR
    IF nPasan = (ULTIMO_PASO + 1) THEN
        veredicto := 1;
    ELSE
        veredicto := 2;
    END_IF
END_IF
